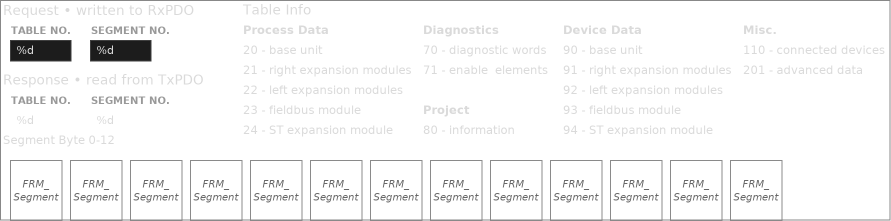
VISUALIZATION FRM_SegmentTable  // 891x221
VAR_IN_OUT
    nRequestTableNo: BYTE;
    nRequestSegmentNo: BYTE;
    
    nResponseTableNo: BYTE;
    nResponseSegmentNo: BYTE;
    
    aSegmentBytes: ARRAY [1..13] OF BYTE;
END_VAR
    Label (0,0 211x21), "Request • written to RxPDO"
    Label (0,70 221x20), "Response • read from TxPDO"
    Textfield (10,110 61x21), "%d", text variable: nResponseTableNo
    Label (8,20 61x21), "TABLE NO."
    Label (88,20 81x21), "SEGMENT NO."
    Textfield (10,40 61x21), "%d", text variable: nRequestTableNo
        OnMouseClick: write the text variable via Default, min 0, max 255
    Textfield (90,40 61x21), "%d", text variable: nRequestSegmentNo
        OnMouseClick: write the text variable via Default, min 0, max 255
    Label (8,90 61x21), "TABLE NO."
    Label (88,90 81x21), "SEGMENT NO."
    Textfield (90,110 61x21), "%d", text variable: nResponseSegmentNo
    Label (0,130 121x20), "Segment Byte 0-12"
    Frame (10,160 52x61)
        shows FRM_Segment(nValue := aSegmentBytes[1], nIndex := 0)
    Frame (70,160 52x61)
        shows FRM_Segment(nValue := aSegmentBytes[2], nIndex := 1)
    Frame (130,160 52x61)
        shows FRM_Segment(nValue := aSegmentBytes[3], nIndex := 2)
    Frame (190,160 52x61)
        shows FRM_Segment(nValue := aSegmentBytes[4], nIndex := 3)
    Frame (250,160 52x61)
        shows FRM_Segment(nValue := aSegmentBytes[5], nIndex := 4)
    Frame (310,160 52x61)
        shows FRM_Segment(nValue := aSegmentBytes[6], nIndex := 5)
    Frame (370,160 52x61)
        shows FRM_Segment(nValue := aSegmentBytes[7], nIndex := 6)
    Frame (430,160 52x61)
        shows FRM_Segment(nValue := aSegmentBytes[8], nIndex := 7)
    Frame (490,160 52x61)
        shows FRM_Segment(nValue := aSegmentBytes[9], nIndex := 8)
    Frame (550,160 52x61)
        shows FRM_Segment(nValue := aSegmentBytes[10], nIndex := 9)
    Frame (610,160 52x61)
        shows FRM_Segment(nValue := aSegmentBytes[11], nIndex := 10)
    Frame (670,160 52x61)
        shows FRM_Segment(nValue := aSegmentBytes[12], nIndex := 11)
    Frame (730,160 52x61)
        shows FRM_Segment(nValue := aSegmentBytes[13], nIndex := 12)
    Label (240,0 81x20), "Table Info"
    Label (240,20 181x20), "Process Data"
    Label (240,40 181x20), "20 - base unit"
    Label (240,60 181x20), "21 - right expansion modules"
    Label (240,80 181x20), "22 - left expansion modules"
    Label (240,100 181x20), "23 - fieldbus module"
    Label (240,120 181x20), "24 - ST expansion module"
    Label (420,20 131x20), "Diagnostics"
    Label (420,40 131x20), "70 - diagnostic words"
    Label (420,60 131x20), "71 - enable elements"
    Label (420,100 131x20), "Project"
    Label (420,120 131x20), "80 - information"
    Label (560,20 181x20), "Device Data"
    Label (560,40 181x20), "90 - base unit"
    Label (560,60 181x20), "91 - right expansion modules"
    Label (560,80 181x20), "92 - left expansion modules"
    Label (560,100 181x20), "93 - fieldbus module"
    Label (560,120 181x20), "94 - ST expansion module"
    Label (740,20 131x20), "Misc."
    Label (740,40 151x20), "110 - connected devices"
    Label (740,60 131x20), "201 - advanced data"
END_VISUALIZATION

(* stored: Version 1.1.0.1
   Visu FRM_SegmentTable: Id {d5754331-7178-0761-3889-f1e808cfc14b} *)
